// Mitsubishi GX Works2 project: TRANG TRAI   PLC: FX3U/FX3UC

PROGRAM MAIN
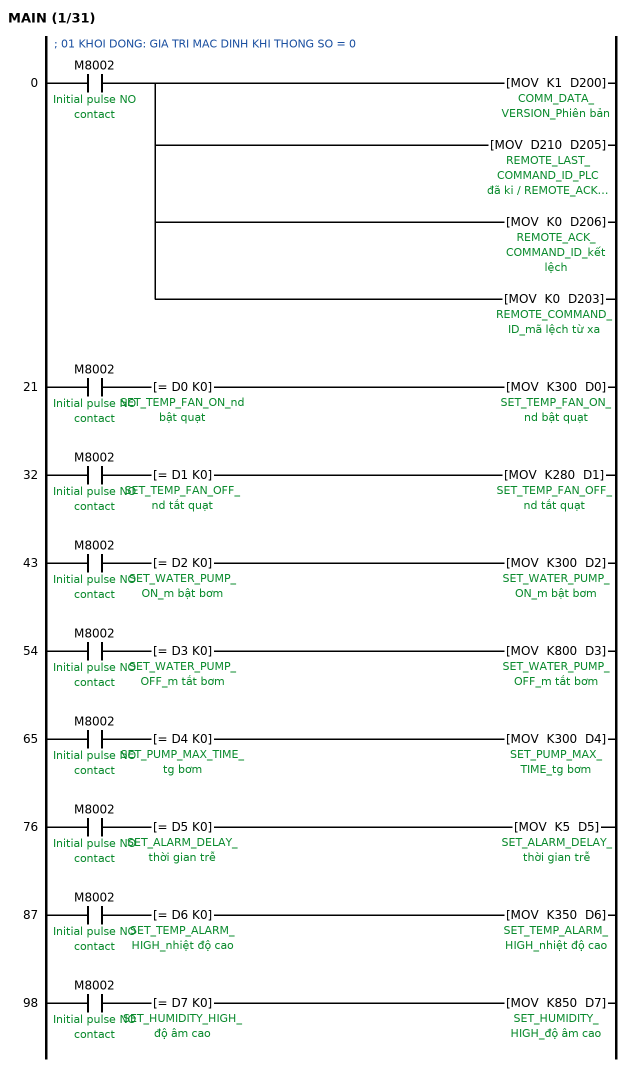
; 01 KHOI DONG: GIA TRI MAC DINH KHI THONG SO = 0
0     LD      M8002  ; Initial pulse NO contact
      MOV     K1 D200  ; COMM_DATA_VERSION_Phiên bản
      MOV     D210 D205  ; REMOTE_LAST_COMMAND_ID_PLC đã ki / REMOTE_ACK_COMMAND_ID_PLC đã nhậ
      MOV     K0 D206  ; REMOTE_ACK_COMMAND_ID_kết lệch
      MOV     K0 D203  ; REMOTE_COMMAND_ID_mã lệch từ xa
21    LD      M8002  ; Initial pulse NO contact
      AND=    D0 K0  ; SET_TEMP_FAN_ON_nd bật quạt
      MOV     K300 D0
32    LD      M8002  ; Initial pulse NO contact
      AND=    D1 K0  ; SET_TEMP_FAN_OFF_nd tắt quạt
      MOV     K280 D1
43    LD      M8002  ; Initial pulse NO contact
      AND=    D2 K0  ; SET_WATER_PUMP_ON_m bật bơm
      MOV     K300 D2
54    LD      M8002  ; Initial pulse NO contact
      AND=    D3 K0  ; SET_WATER_PUMP_OFF_m tắt bơm
      MOV     K800 D3
65    LD      M8002  ; Initial pulse NO contact
      AND=    D4 K0  ; SET_PUMP_MAX_TIME_tg bơm
      MOV     K300 D4
76    LD      M8002  ; Initial pulse NO contact
      AND=    D5 K0  ; SET_ALARM_DELAY_thời gian trễ
      MOV     K5 D5
87    LD      M8002  ; Initial pulse NO contact
      AND=    D6 K0  ; SET_TEMP_ALARM_HIGH_nhiệt độ cao
      MOV     K350 D6
98    LD      M8002  ; Initial pulse NO contact
      AND=    D7 K0  ; SET_HUMIDITY_HIGH_độ âm cao
      MOV     K850 D7
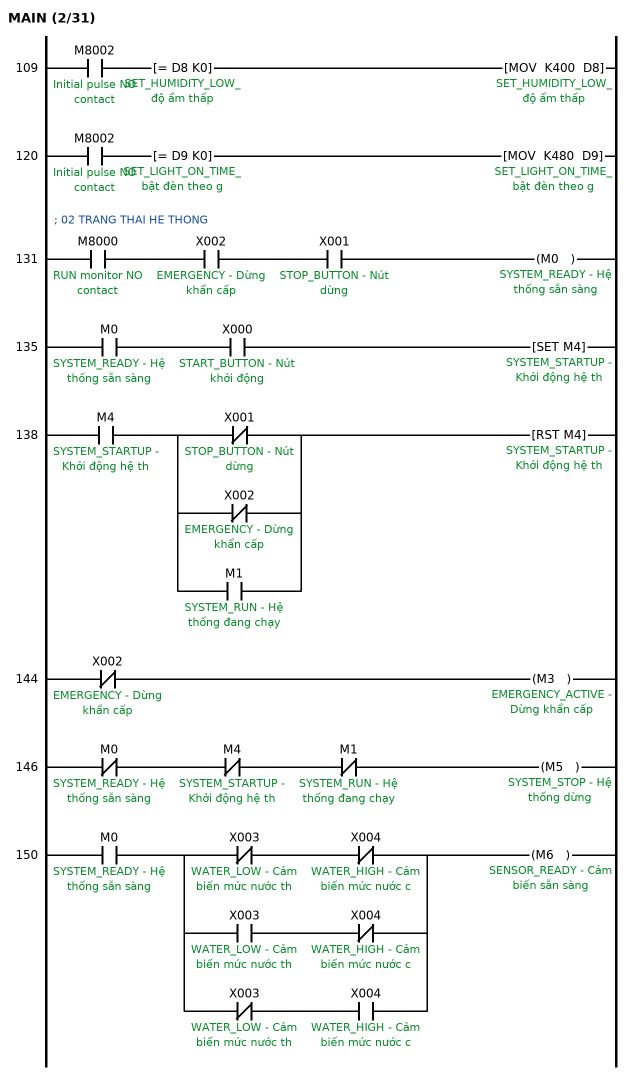
109   LD      M8002  ; Initial pulse NO contact
      AND=    D8 K0  ; SET_HUMIDITY_LOW_độ ẩm thấp
      MOV     K400 D8
120   LD      M8002  ; Initial pulse NO contact
      AND=    D9 K0  ; SET_LIGHT_ON_TIME_bật đèn theo g
      MOV     K480 D9
; 02 TRANG THAI HE THONG
131   LD      M8000  ; RUN monitor NO contact
      AND     X002  ; EMERGENCY - Dừng khẩn cấp
      AND     X001  ; STOP_BUTTON - Nút dừng
      OUT     M0  ; SYSTEM_READY - Hệ thống sẵn sàng
135   LD      M0  ; SYSTEM_READY - Hệ thống sẵn sàng
      AND     X000  ; START_BUTTON - Nút khởi động
      SET     M4  ; SYSTEM_STARTUP - Khởi động hệ th
138   LD      M4  ; SYSTEM_STARTUP - Khởi động hệ th
      LDI     X001  ; STOP_BUTTON - Nút dừng
      ORI     X002  ; EMERGENCY - Dừng khẩn cấp
      OR      M1  ; SYSTEM_RUN - Hệ thống đang chạy
      ANB
      RST     M4  ; SYSTEM_STARTUP - Khởi động hệ th
144   LDI     X002  ; EMERGENCY - Dừng khẩn cấp
      OUT     M3  ; EMERGENCY_ACTIVE - Dừng khẩn cấp
146   LDI     M0  ; SYSTEM_READY - Hệ thống sẵn sàng
      ANI     M4  ; SYSTEM_STARTUP - Khởi động hệ th
      ANI     M1  ; SYSTEM_RUN - Hệ thống đang chạy
      OUT     M5  ; SYSTEM_STOP - Hệ thống dừng
150   LD      M0  ; SYSTEM_READY - Hệ thống sẵn sàng
      LDI     X003  ; WATER_LOW - Cảm biến mức nước th
      ANI     X004  ; WATER_HIGH - Cảm biến mức nước c
      LD      X003  ; WATER_LOW - Cảm biến mức nước th
      ANI     X004  ; WATER_HIGH - Cảm biến mức nước c
      ORB
      LDI     X003  ; WATER_LOW - Cảm biến mức nước th
      AND     X004  ; WATER_HIGH - Cảm biến mức nước c
      ORB
      ANB
      OUT     M6  ; SENSOR_READY - Cảm biến sẵn sàng
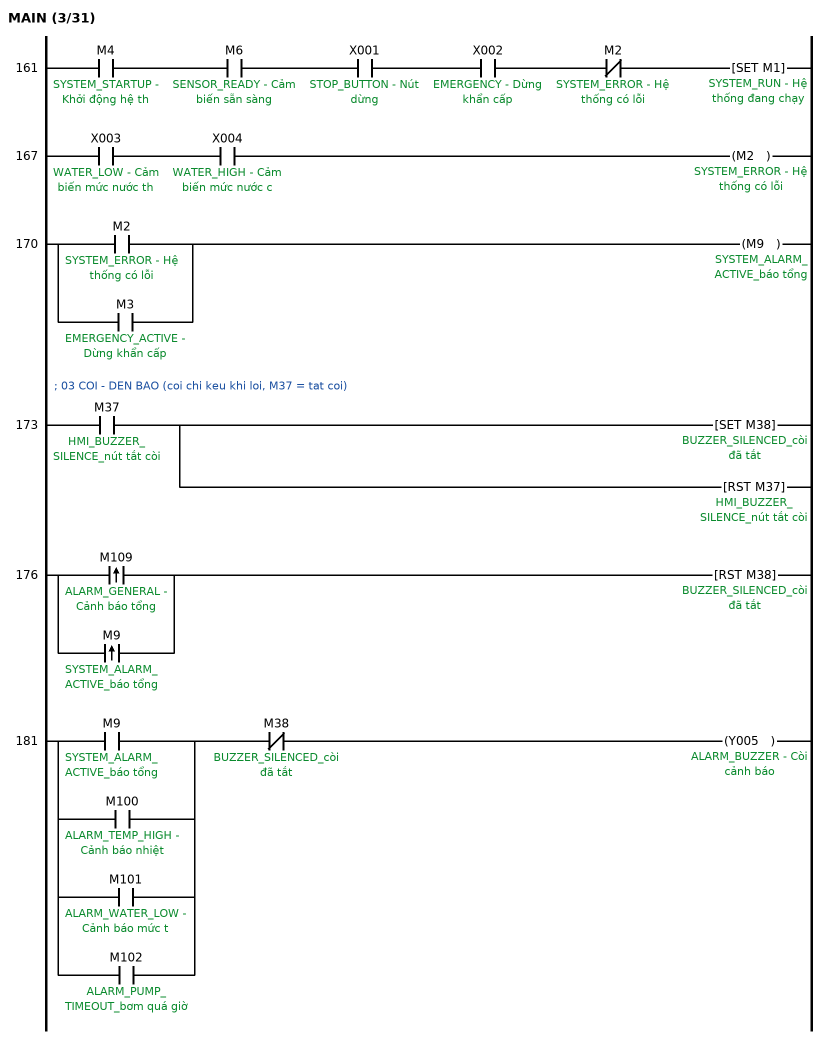
161   LD      M4  ; SYSTEM_STARTUP - Khởi động hệ th
      AND     M6  ; SENSOR_READY - Cảm biến sẵn sàng
      AND     X001  ; STOP_BUTTON - Nút dừng
      AND     X002  ; EMERGENCY - Dừng khẩn cấp
      ANI     M2  ; SYSTEM_ERROR - Hệ thống có lỗi
      SET     M1  ; SYSTEM_RUN - Hệ thống đang chạy
167   LD      X003  ; WATER_LOW - Cảm biến mức nước th
      AND     X004  ; WATER_HIGH - Cảm biến mức nước c
      OUT     M2  ; SYSTEM_ERROR - Hệ thống có lỗi
170   LD      M2  ; SYSTEM_ERROR - Hệ thống có lỗi
      OR      M3  ; EMERGENCY_ACTIVE - Dừng khẩn cấp
      OUT     M9  ; SYSTEM_ALARM_ACTIVE_báo tổng
; 03 COI - DEN BAO (coi chi keu khi loi, M37 = tat coi)
173   LD      M37  ; HMI_BUZZER_SILENCE_nút tắt còi
      SET     M38  ; BUZZER_SILENCED_còi đã tắt
      RST     M37  ; HMI_BUZZER_SILENCE_nút tắt còi
176   LDP     M109  ; ALARM_GENERAL - Cảnh báo tổng
      ORP     M9  ; SYSTEM_ALARM_ACTIVE_báo tổng
      RST     M38  ; BUZZER_SILENCED_còi đã tắt
181   LD      M9  ; SYSTEM_ALARM_ACTIVE_báo tổng
      OR      M100  ; ALARM_TEMP_HIGH - Cảnh báo nhiệt
      OR      M101  ; ALARM_WATER_LOW - Cảnh báo mức t
      OR      M102  ; ALARM_PUMP_TIMEOUT_bơm quá giờ
      ANI     M38  ; BUZZER_SILENCED_còi đã tắt
      OUT     Y005  ; ALARM_BUZZER - Còi cảnh báo
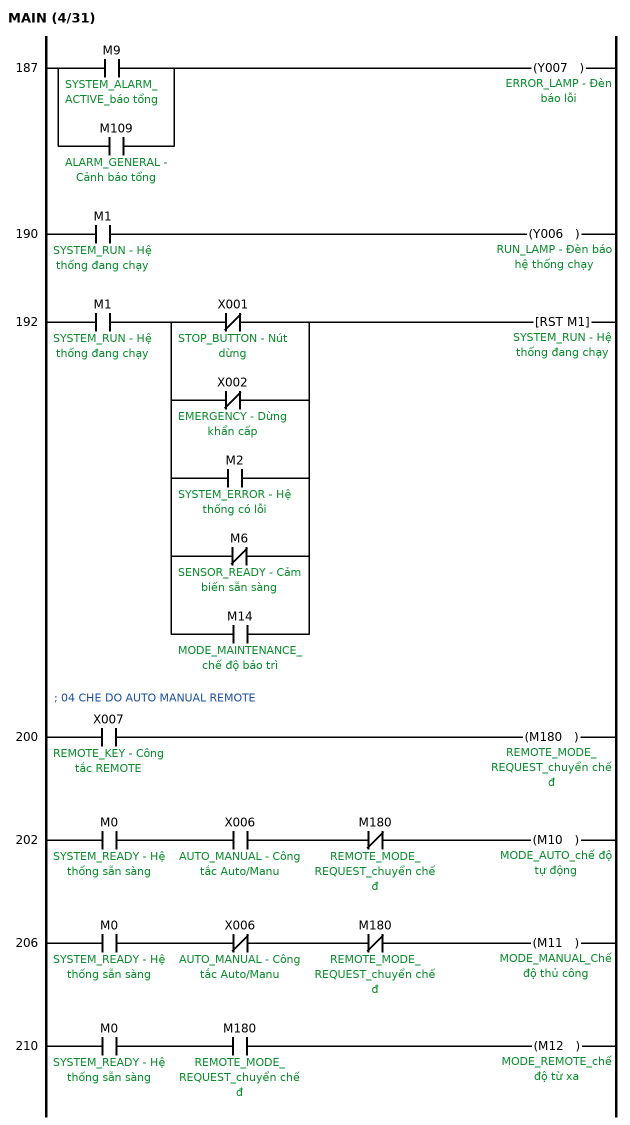
187   LD      M9  ; SYSTEM_ALARM_ACTIVE_báo tổng
      OR      M109  ; ALARM_GENERAL - Cảnh báo tổng
      OUT     Y007  ; ERROR_LAMP - Đèn báo lỗi
190   LD      M1  ; SYSTEM_RUN - Hệ thống đang chạy
      OUT     Y006  ; RUN_LAMP - Đèn báo hệ thống chạy
192   LD      M1  ; SYSTEM_RUN - Hệ thống đang chạy
      LDI     X001  ; STOP_BUTTON - Nút dừng
      ORI     X002  ; EMERGENCY - Dừng khẩn cấp
      OR      M2  ; SYSTEM_ERROR - Hệ thống có lỗi
      ORI     M6  ; SENSOR_READY - Cảm biến sẵn sàng
      OR      M14  ; MODE_MAINTENANCE_chế độ bảo trì
      ANB
      RST     M1  ; SYSTEM_RUN - Hệ thống đang chạy
; 04 CHE DO AUTO MANUAL REMOTE
200   LD      X007  ; REMOTE_KEY - Công tắc REMOTE
      OUT     M180  ; REMOTE_MODE_REQUEST_chuyển chế đ
202   LD      M0  ; SYSTEM_READY - Hệ thống sẵn sàng
      AND     X006  ; AUTO_MANUAL - Công tắc Auto/Manu
      ANI     M180  ; REMOTE_MODE_REQUEST_chuyển chế đ
      OUT     M10  ; MODE_AUTO_chế độ tự động
206   LD      M0  ; SYSTEM_READY - Hệ thống sẵn sàng
      ANI     X006  ; AUTO_MANUAL - Công tắc Auto/Manu
      ANI     M180  ; REMOTE_MODE_REQUEST_chuyển chế đ
      OUT     M11  ; MODE_MANUAL_Chế độ thủ công
210   LD      M0  ; SYSTEM_READY - Hệ thống sẵn sàng
      AND     M180  ; REMOTE_MODE_REQUEST_chuyển chế đ
      OUT     M12  ; MODE_REMOTE_chế độ từ xa
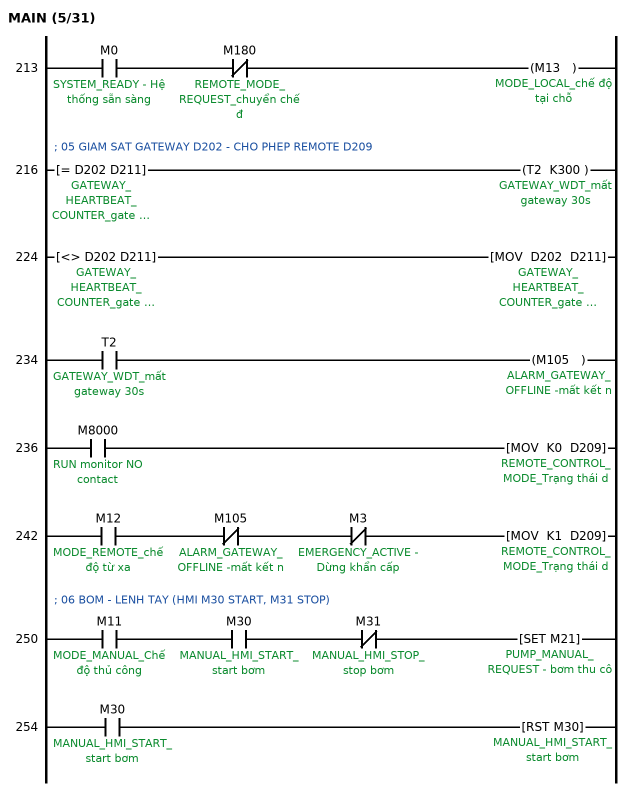
213   LD      M0  ; SYSTEM_READY - Hệ thống sẵn sàng
      ANI     M180  ; REMOTE_MODE_REQUEST_chuyển chế đ
      OUT     M13  ; MODE_LOCAL_chế độ tại chỗ
; 05 GIAM SAT GATEWAY D202 - CHO PHEP REMOTE D209
216   LD=     D202 D211  ; GATEWAY_HEARTBEAT_COUNTER_gate / GATEWAY_HB_LAST_D202 lần trước
      OUT     T2 K300  ; GATEWAY_WDT_mất gateway 30s
224   LD<>    D202 D211  ; GATEWAY_HEARTBEAT_COUNTER_gate / GATEWAY_HB_LAST_D202 lần trước
      MOV     D202 D211
234   LD      T2  ; GATEWAY_WDT_mất gateway 30s
      OUT     M105  ; ALARM_GATEWAY_OFFLINE -mất kết n
236   LD      M8000  ; RUN monitor NO contact
      MOV     K0 D209  ; REMOTE_CONTROL_MODE_Trạng thái d
242   LD      M12  ; MODE_REMOTE_chế độ từ xa
      ANI     M105  ; ALARM_GATEWAY_OFFLINE -mất kết n
      ANI     M3  ; EMERGENCY_ACTIVE - Dừng khẩn cấp
      MOV     K1 D209
; 06 BOM - LENH TAY (HMI M30 START, M31 STOP)
250   LD      M11  ; MODE_MANUAL_Chế độ thủ công
      AND     M30  ; MANUAL_HMI_START_start bơm
      ANI     M31  ; MANUAL_HMI_STOP_stop bơm
      SET     M21  ; PUMP_MANUAL_REQUEST - bơm thu cô
254   LD      M30  ; MANUAL_HMI_START_start bơm
      RST     M30  ; MANUAL_HMI_START_start bơm
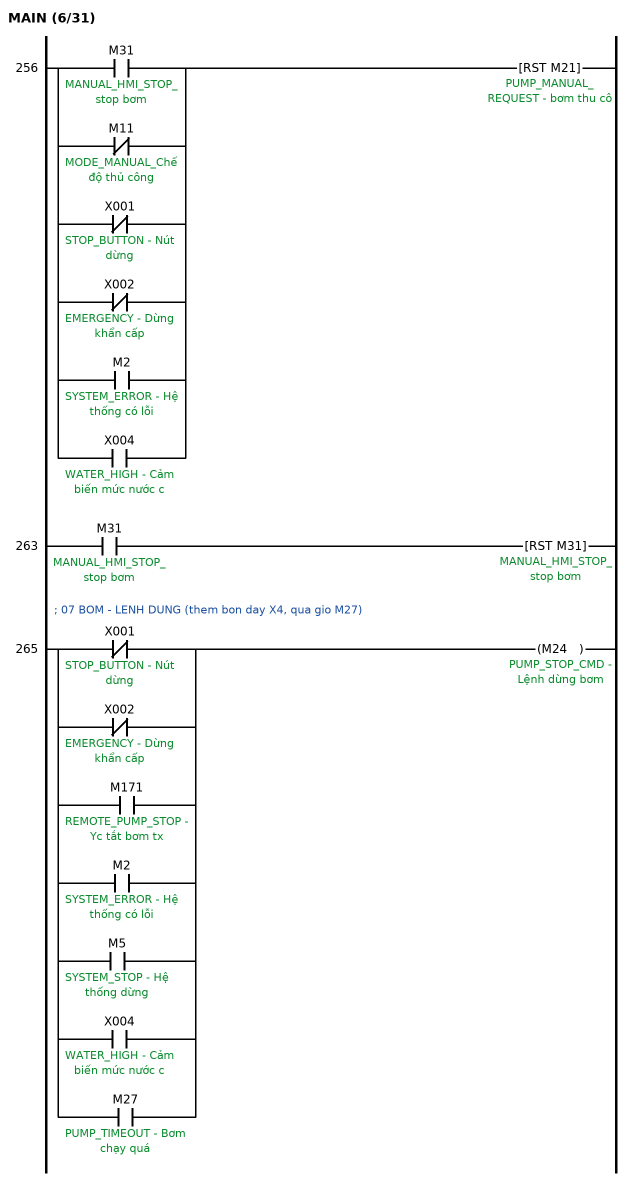
256   LD      M31  ; MANUAL_HMI_STOP_stop bơm
      ORI     M11  ; MODE_MANUAL_Chế độ thủ công
      ORI     X001  ; STOP_BUTTON - Nút dừng
      ORI     X002  ; EMERGENCY - Dừng khẩn cấp
      OR      M2  ; SYSTEM_ERROR - Hệ thống có lỗi
      OR      X004  ; WATER_HIGH - Cảm biến mức nước c
      RST     M21  ; PUMP_MANUAL_REQUEST - bơm thu cô
263   LD      M31  ; MANUAL_HMI_STOP_stop bơm
      RST     M31  ; MANUAL_HMI_STOP_stop bơm
; 07 BOM - LENH DUNG (them bon day X4, qua gio M27)
265   LDI     X001  ; STOP_BUTTON - Nút dừng
      ORI     X002  ; EMERGENCY - Dừng khẩn cấp
      OR      M171  ; REMOTE_PUMP_STOP - Yc tắt bơm tx
      OR      M2  ; SYSTEM_ERROR - Hệ thống có lỗi
      OR      M5  ; SYSTEM_STOP - Hệ thống dừng
      OR      X004  ; WATER_HIGH - Cảm biến mức nước c
      OR      M27  ; PUMP_TIMEOUT - Bơm chạy quá
      OUT     M24  ; PUMP_STOP_CMD - Lệnh dừng bơm
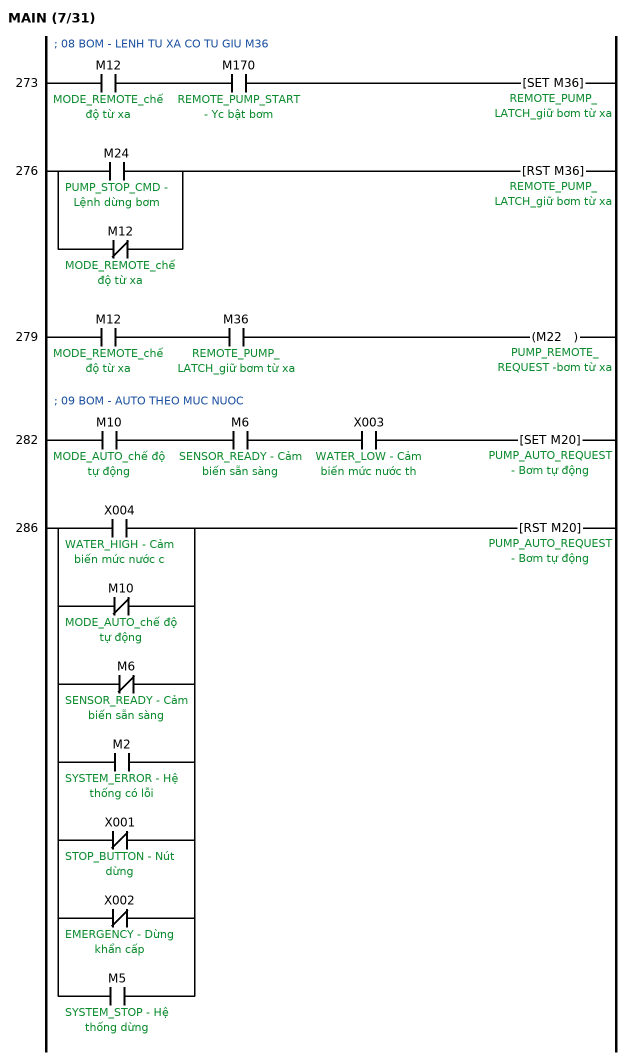
; 08 BOM - LENH TU XA CO TU GIU M36
273   LD      M12  ; MODE_REMOTE_chế độ từ xa
      AND     M170  ; REMOTE_PUMP_START - Yc bật bơm
      SET     M36  ; REMOTE_PUMP_LATCH_giữ bơm từ xa
276   LD      M24  ; PUMP_STOP_CMD - Lệnh dừng bơm
      ORI     M12  ; MODE_REMOTE_chế độ từ xa
      RST     M36  ; REMOTE_PUMP_LATCH_giữ bơm từ xa
279   LD      M12  ; MODE_REMOTE_chế độ từ xa
      AND     M36  ; REMOTE_PUMP_LATCH_giữ bơm từ xa
      OUT     M22  ; PUMP_REMOTE_REQUEST -bơm từ xa
; 09 BOM - AUTO THEO MUC NUOC
282   LD      M10  ; MODE_AUTO_chế độ tự động
      AND     M6  ; SENSOR_READY - Cảm biến sẵn sàng
      AND     X003  ; WATER_LOW - Cảm biến mức nước th
      SET     M20  ; PUMP_AUTO_REQUEST - Bơm tự động
286   LD      X004  ; WATER_HIGH - Cảm biến mức nước c
      ORI     M10  ; MODE_AUTO_chế độ tự động
      ORI     M6  ; SENSOR_READY - Cảm biến sẵn sàng
      OR      M2  ; SYSTEM_ERROR - Hệ thống có lỗi
      ORI     X001  ; STOP_BUTTON - Nút dừng
      ORI     X002  ; EMERGENCY - Dừng khẩn cấp
      OR      M5  ; SYSTEM_STOP - Hệ thống dừng
      RST     M20  ; PUMP_AUTO_REQUEST - Bơm tự động
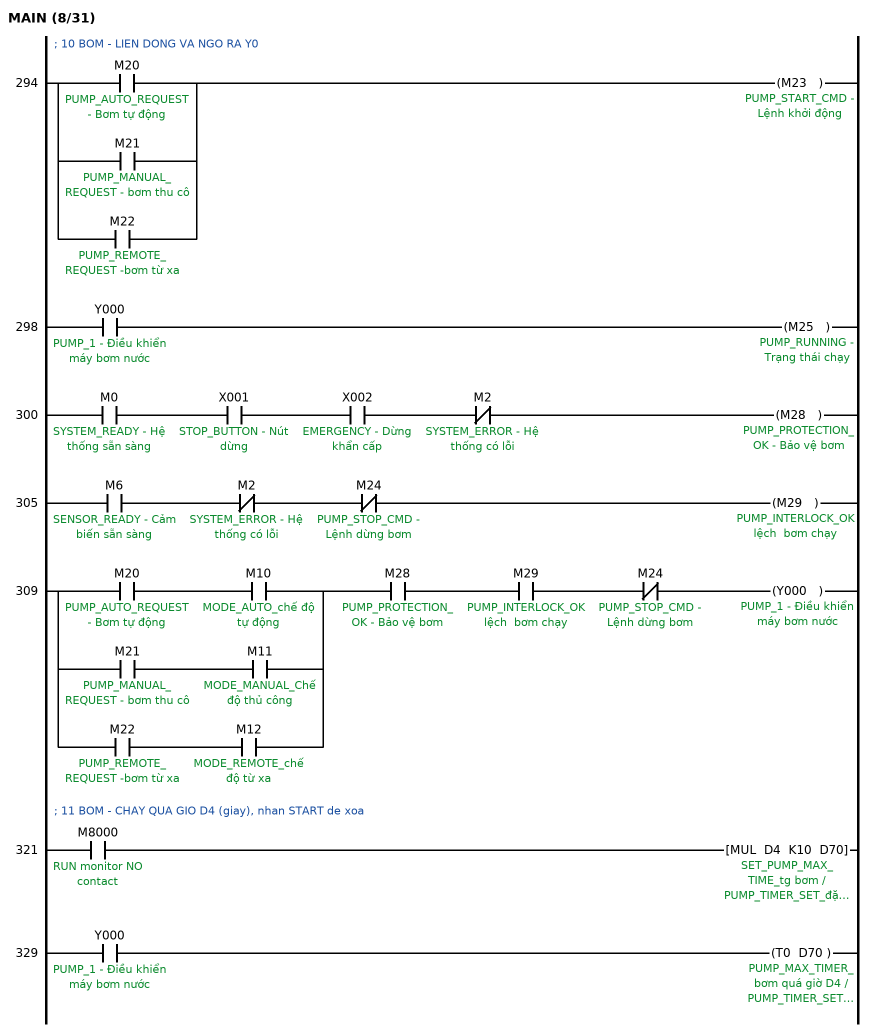
; 10 BOM - LIEN DONG VA NGO RA Y0
294   LD      M20  ; PUMP_AUTO_REQUEST - Bơm tự động
      OR      M21  ; PUMP_MANUAL_REQUEST - bơm thu cô
      OR      M22  ; PUMP_REMOTE_REQUEST -bơm từ xa
      OUT     M23  ; PUMP_START_CMD - Lệnh khởi động
298   LD      Y000  ; PUMP_1 - Điều khiển máy bơm nước
      OUT     M25  ; PUMP_RUNNING - Trạng thái chạy
300   LD      M0  ; SYSTEM_READY - Hệ thống sẵn sàng
      AND     X001  ; STOP_BUTTON - Nút dừng
      AND     X002  ; EMERGENCY - Dừng khẩn cấp
      ANI     M2  ; SYSTEM_ERROR - Hệ thống có lỗi
      OUT     M28  ; PUMP_PROTECTION_OK - Bảo vệ bơm
305   LD      M6  ; SENSOR_READY - Cảm biến sẵn sàng
      ANI     M2  ; SYSTEM_ERROR - Hệ thống có lỗi
      ANI     M24  ; PUMP_STOP_CMD - Lệnh dừng bơm
      OUT     M29  ; PUMP_INTERLOCK_OK lệch  bơm chạy
309   LD      M20  ; PUMP_AUTO_REQUEST - Bơm tự động
      AND     M10  ; MODE_AUTO_chế độ tự động
      LD      M21  ; PUMP_MANUAL_REQUEST - bơm thu cô
      AND     M11  ; MODE_MANUAL_Chế độ thủ công
      ORB
      LD      M22  ; PUMP_REMOTE_REQUEST -bơm từ xa
      AND     M12  ; MODE_REMOTE_chế độ từ xa
      ORB
      AND     M28  ; PUMP_PROTECTION_OK - Bảo vệ bơm
      AND     M29  ; PUMP_INTERLOCK_OK lệch  bơm chạy
      ANI     M24  ; PUMP_STOP_CMD - Lệnh dừng bơm
      OUT     Y000  ; PUMP_1 - Điều khiển máy bơm nước
; 11 BOM - CHAY QUA GIO D4 (giay), nhan START de xoa
321   LD      M8000  ; RUN monitor NO contact
      MUL     D4 K10 D70  ; PUMP_TIMER_SET_đặt T0 = D4x10
329   LD      Y000  ; PUMP_1 - Điều khiển máy bơm nước
      OUT     T0 D70  ; PUMP_MAX_TIMER_bơm quá giờ D4 / PUMP_TIMER_SET_đặt T0 = D4x10
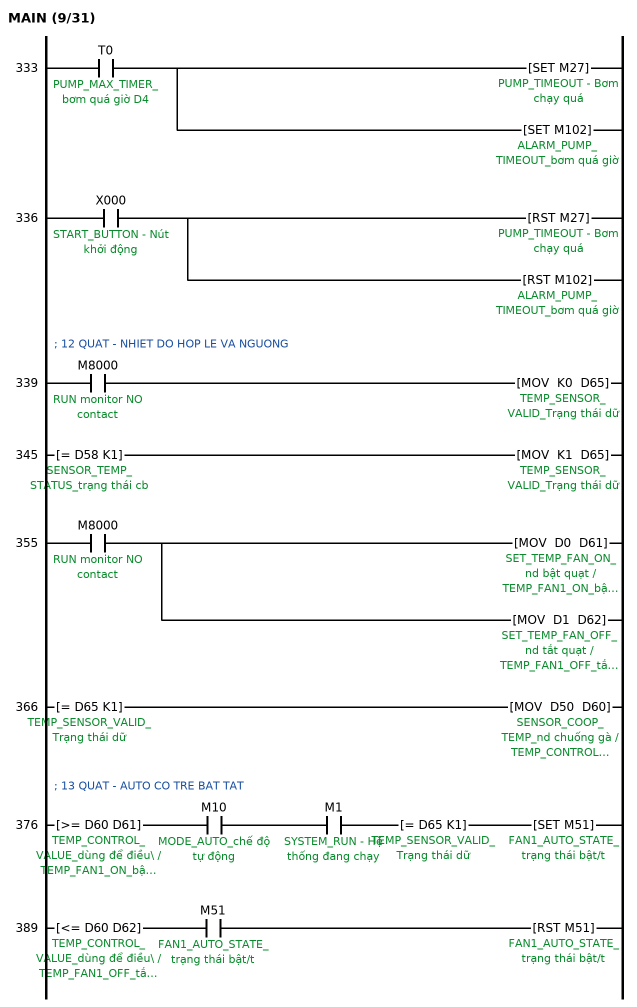
333   LD      T0  ; PUMP_MAX_TIMER_bơm quá giờ D4
      SET     M27  ; PUMP_TIMEOUT - Bơm chạy quá
      SET     M102  ; ALARM_PUMP_TIMEOUT_bơm quá giờ
336   LD      X000  ; START_BUTTON - Nút khởi động
      RST     M27  ; PUMP_TIMEOUT - Bơm chạy quá
      RST     M102  ; ALARM_PUMP_TIMEOUT_bơm quá giờ
; 12 QUAT - NHIET DO HOP LE VA NGUONG
339   LD      M8000  ; RUN monitor NO contact
      MOV     K0 D65  ; TEMP_SENSOR_VALID_Trạng thái dữ
345   LD=     D58 K1  ; SENSOR_TEMP_STATUS_trạng thái cb
      MOV     K1 D65
355   LD      M8000  ; RUN monitor NO contact
      MOV     D0 D61  ; TEMP_FAN1_ON_bật quạt 1
      MOV     D1 D62  ; TEMP_FAN1_OFF_tắt quạt 1
366   LD=     D65 K1  ; TEMP_SENSOR_VALID_Trạng thái dữ
      MOV     D50 D60  ; SENSOR_COOP_TEMP_nd chuống gà / TEMP_CONTROL_VALUE_dùng để điều\
; 13 QUAT - AUTO CO TRE BAT TAT
376   LD>=    D60 D61  ; TEMP_CONTROL_VALUE_dùng để điều\ / TEMP_FAN1_ON_bật quạt 1
      AND     M10  ; MODE_AUTO_chế độ tự động
      AND     M1  ; SYSTEM_RUN - Hệ thống đang chạy
      AND=    D65 K1  ; TEMP_SENSOR_VALID_Trạng thái dữ
      SET     M51  ; FAN1_AUTO_STATE_trạng thái bật/t
389   LD<=    D60 D62  ; TEMP_CONTROL_VALUE_dùng để điều\ / TEMP_FAN1_OFF_tắt quạt 1
      AND     M51  ; FAN1_AUTO_STATE_trạng thái bật/t
      RST     M51  ; FAN1_AUTO_STATE_trạng thái bật/t
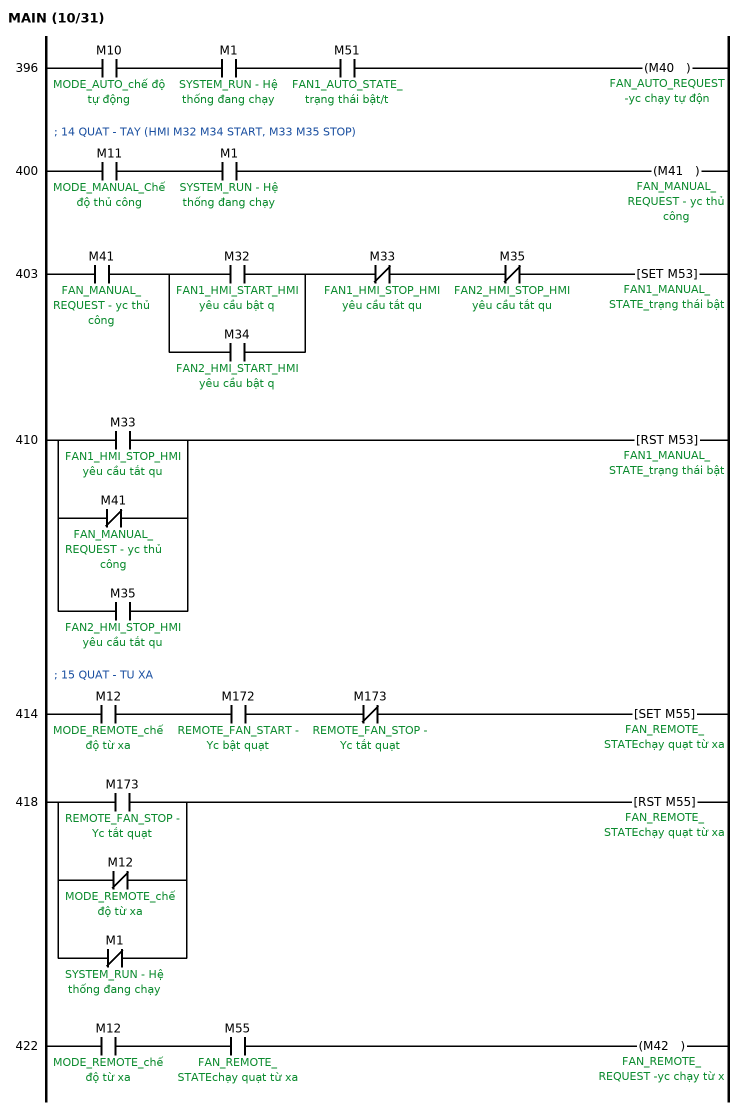
396   LD      M10  ; MODE_AUTO_chế độ tự động
      AND     M1  ; SYSTEM_RUN - Hệ thống đang chạy
      AND     M51  ; FAN1_AUTO_STATE_trạng thái bật/t
      OUT     M40  ; FAN_AUTO_REQUEST -yc chạy tự độn
; 14 QUAT - TAY (HMI M32 M34 START, M33 M35 STOP)
400   LD      M11  ; MODE_MANUAL_Chế độ thủ công
      AND     M1  ; SYSTEM_RUN - Hệ thống đang chạy
      OUT     M41  ; FAN_MANUAL_REQUEST - yc thủ công
403   LD      M41  ; FAN_MANUAL_REQUEST - yc thủ công
      LD      M32  ; FAN1_HMI_START_HMI yêu cầu bật q
      OR      M34  ; FAN2_HMI_START_HMI yêu cầu bật q
      ANB
      ANI     M33  ; FAN1_HMI_STOP_HMI yêu cầu tắt qu
      ANI     M35  ; FAN2_HMI_STOP_HMI yêu cầu tắt qu
      SET     M53  ; FAN1_MANUAL_STATE_trạng thái bật
410   LD      M33  ; FAN1_HMI_STOP_HMI yêu cầu tắt qu
      ORI     M41  ; FAN_MANUAL_REQUEST - yc thủ công
      OR      M35  ; FAN2_HMI_STOP_HMI yêu cầu tắt qu
      RST     M53  ; FAN1_MANUAL_STATE_trạng thái bật
; 15 QUAT - TU XA
414   LD      M12  ; MODE_REMOTE_chế độ từ xa
      AND     M172  ; REMOTE_FAN_START - Yc bật quạt
      ANI     M173  ; REMOTE_FAN_STOP - Yc tắt quạt
      SET     M55  ; FAN_REMOTE_STATEchạy quạt từ xa
418   LD      M173  ; REMOTE_FAN_STOP - Yc tắt quạt
      ORI     M12  ; MODE_REMOTE_chế độ từ xa
      ORI     M1  ; SYSTEM_RUN - Hệ thống đang chạy
      RST     M55  ; FAN_REMOTE_STATEchạy quạt từ xa
422   LD      M12  ; MODE_REMOTE_chế độ từ xa
      AND     M55  ; FAN_REMOTE_STATEchạy quạt từ xa
      OUT     M42  ; FAN_REMOTE_REQUEST -yc chạy từ x
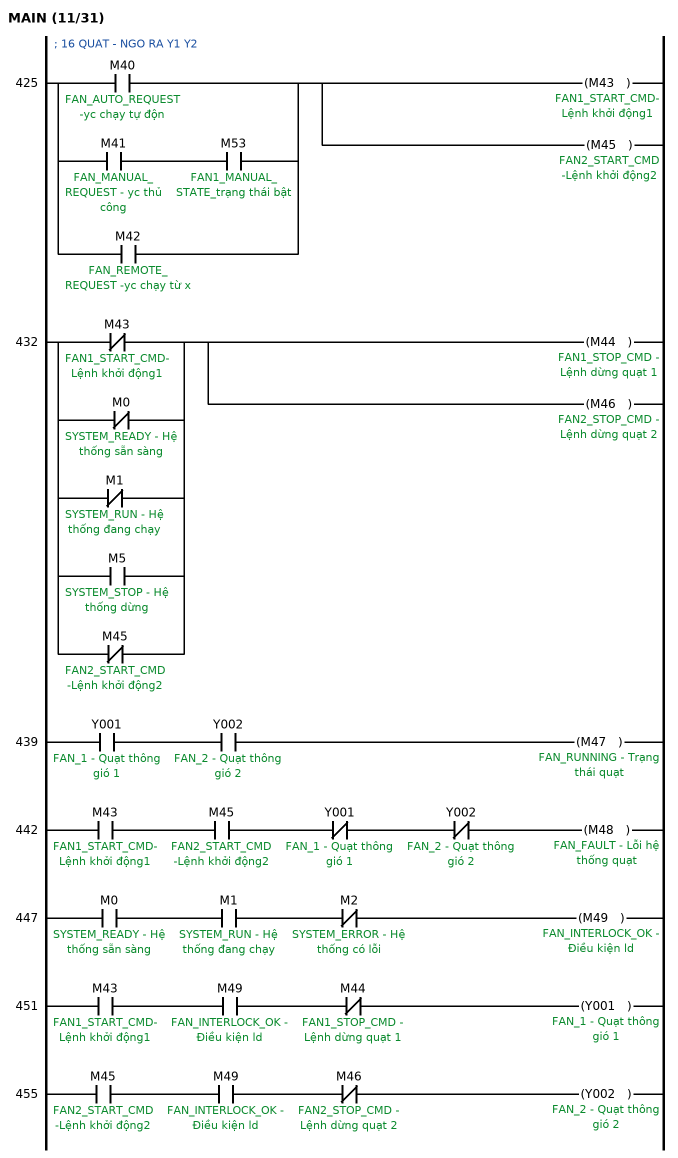
; 16 QUAT - NGO RA Y1 Y2
425   LD      M40  ; FAN_AUTO_REQUEST -yc chạy tự độn
      LD      M41  ; FAN_MANUAL_REQUEST - yc thủ công
      AND     M53  ; FAN1_MANUAL_STATE_trạng thái bật
      ORB
      OR      M42  ; FAN_REMOTE_REQUEST -yc chạy từ x
      OUT     M43  ; FAN1_START_CMD-Lệnh khởi động1
      OUT     M45  ; FAN2_START_CMD -Lệnh khởi động2
432   LDI     M43  ; FAN1_START_CMD-Lệnh khởi động1
      ORI     M0  ; SYSTEM_READY - Hệ thống sẵn sàng
      ORI     M1  ; SYSTEM_RUN - Hệ thống đang chạy
      OR      M5  ; SYSTEM_STOP - Hệ thống dừng
      ORI     M45  ; FAN2_START_CMD -Lệnh khởi động2
      OUT     M44  ; FAN1_STOP_CMD - Lệnh dừng quạt 1
      OUT     M46  ; FAN2_STOP_CMD - Lệnh dừng quạt 2
439   LD      Y001  ; FAN_1 - Quạt thông gió 1
      AND     Y002  ; FAN_2 - Quạt thông gió 2
      OUT     M47  ; FAN_RUNNING - Trạng thái quạt
442   LD      M43  ; FAN1_START_CMD-Lệnh khởi động1
      AND     M45  ; FAN2_START_CMD -Lệnh khởi động2
      ANI     Y001  ; FAN_1 - Quạt thông gió 1
      ANI     Y002  ; FAN_2 - Quạt thông gió 2
      OUT     M48  ; FAN_FAULT - Lỗi hệ thống quạt
447   LD      M0  ; SYSTEM_READY - Hệ thống sẵn sàng
      AND     M1  ; SYSTEM_RUN - Hệ thống đang chạy
      ANI     M2  ; SYSTEM_ERROR - Hệ thống có lỗi
      OUT     M49  ; FAN_INTERLOCK_OK - Điều kiện ld
451   LD      M43  ; FAN1_START_CMD-Lệnh khởi động1
      AND     M49  ; FAN_INTERLOCK_OK - Điều kiện ld
      ANI     M44  ; FAN1_STOP_CMD - Lệnh dừng quạt 1
      OUT     Y001  ; FAN_1 - Quạt thông gió 1
455   LD      M45  ; FAN2_START_CMD -Lệnh khởi động2
      AND     M49  ; FAN_INTERLOCK_OK - Điều kiện ld
      ANI     M46  ; FAN2_STOP_CMD - Lệnh dừng quạt 2
      OUT     Y002  ; FAN_2 - Quạt thông gió 2
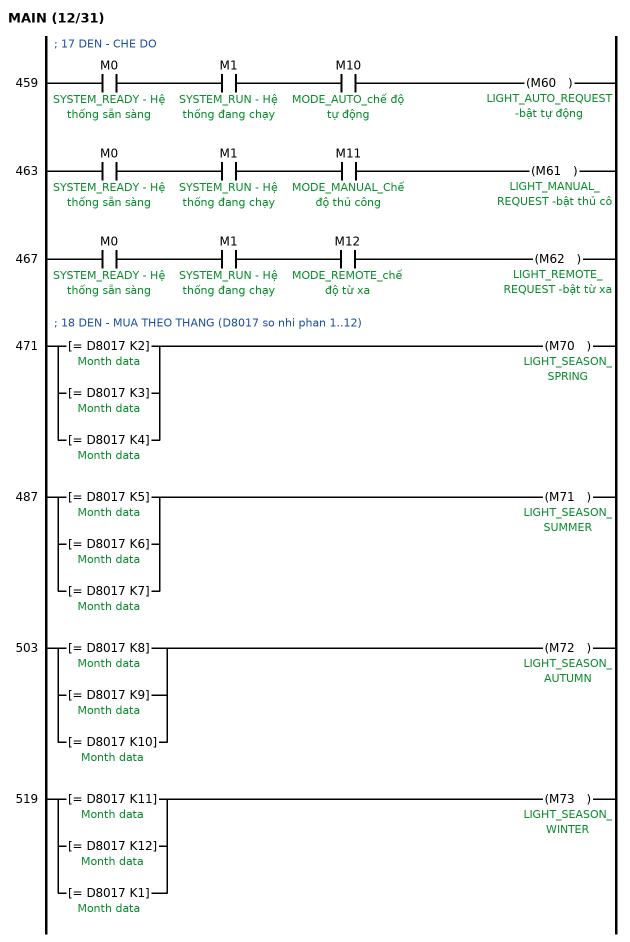
; 17 DEN - CHE DO
459   LD      M0  ; SYSTEM_READY - Hệ thống sẵn sàng
      AND     M1  ; SYSTEM_RUN - Hệ thống đang chạy
      AND     M10  ; MODE_AUTO_chế độ tự động
      OUT     M60  ; LIGHT_AUTO_REQUEST -bật tự động
463   LD      M0  ; SYSTEM_READY - Hệ thống sẵn sàng
      AND     M1  ; SYSTEM_RUN - Hệ thống đang chạy
      AND     M11  ; MODE_MANUAL_Chế độ thủ công
      OUT     M61  ; LIGHT_MANUAL_REQUEST -bật thủ cô
467   LD      M0  ; SYSTEM_READY - Hệ thống sẵn sàng
      AND     M1  ; SYSTEM_RUN - Hệ thống đang chạy
      AND     M12  ; MODE_REMOTE_chế độ từ xa
      OUT     M62  ; LIGHT_REMOTE_REQUEST -bật từ xa
; 18 DEN - MUA THEO THANG (D8017 so nhi phan 1..12)
471   LD=     D8017 K2  ; Month data
      OR=     D8017 K3  ; Month data
      OR=     D8017 K4  ; Month data
      OUT     M70  ; LIGHT_SEASON_SPRING
487   LD=     D8017 K5  ; Month data
      OR=     D8017 K6  ; Month data
      OR=     D8017 K7  ; Month data
      OUT     M71  ; LIGHT_SEASON_SUMMER
503   LD=     D8017 K8  ; Month data
      OR=     D8017 K9  ; Month data
      OR=     D8017 K10  ; Month data
      OUT     M72  ; LIGHT_SEASON_AUTUMN
519   LD=     D8017 K11  ; Month data
      OR=     D8017 K12  ; Month data
      OR=     D8017 K1  ; Month data
      OUT     M73  ; LIGHT_SEASON_WINTER
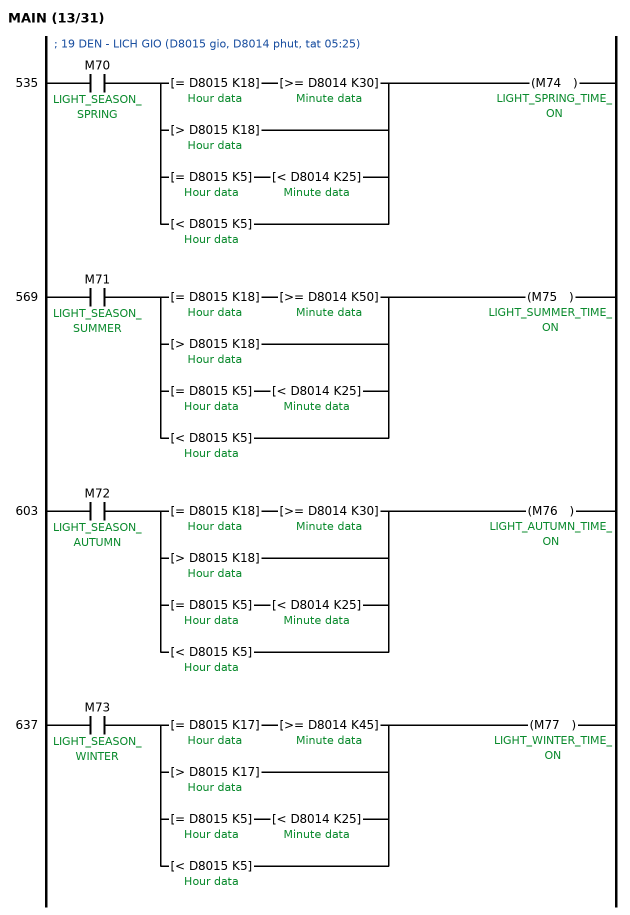
; 19 DEN - LICH GIO (D8015 gio, D8014 phut, tat 05:25)
535   LD      M70  ; LIGHT_SEASON_SPRING
      LD=     D8015 K18  ; Hour data
      AND>=   D8014 K30  ; Minute data
      OR>     D8015 K18  ; Hour data
      LD=     D8015 K5  ; Hour data
      AND<    D8014 K25  ; Minute data
      ORB
      OR<     D8015 K5  ; Hour data
      ANB
      OUT     M74  ; LIGHT_SPRING_TIME_ON
569   LD      M71  ; LIGHT_SEASON_SUMMER
      LD=     D8015 K18  ; Hour data
      AND>=   D8014 K50  ; Minute data
      OR>     D8015 K18  ; Hour data
      LD=     D8015 K5  ; Hour data
      AND<    D8014 K25  ; Minute data
      ORB
      OR<     D8015 K5  ; Hour data
      ANB
      OUT     M75  ; LIGHT_SUMMER_TIME_ON
603   LD      M72  ; LIGHT_SEASON_AUTUMN
      LD=     D8015 K18  ; Hour data
      AND>=   D8014 K30  ; Minute data
      OR>     D8015 K18  ; Hour data
      LD=     D8015 K5  ; Hour data
      AND<    D8014 K25  ; Minute data
      ORB
      OR<     D8015 K5  ; Hour data
      ANB
      OUT     M76  ; LIGHT_AUTUMN_TIME_ON
637   LD      M73  ; LIGHT_SEASON_WINTER
      LD=     D8015 K17  ; Hour data
      AND>=   D8014 K45  ; Minute data
      OR>     D8015 K17  ; Hour data
      LD=     D8015 K5  ; Hour data
      AND<    D8014 K25  ; Minute data
      ORB
      OR<     D8015 K5  ; Hour data
      ANB
      OUT     M77  ; LIGHT_WINTER_TIME_ON
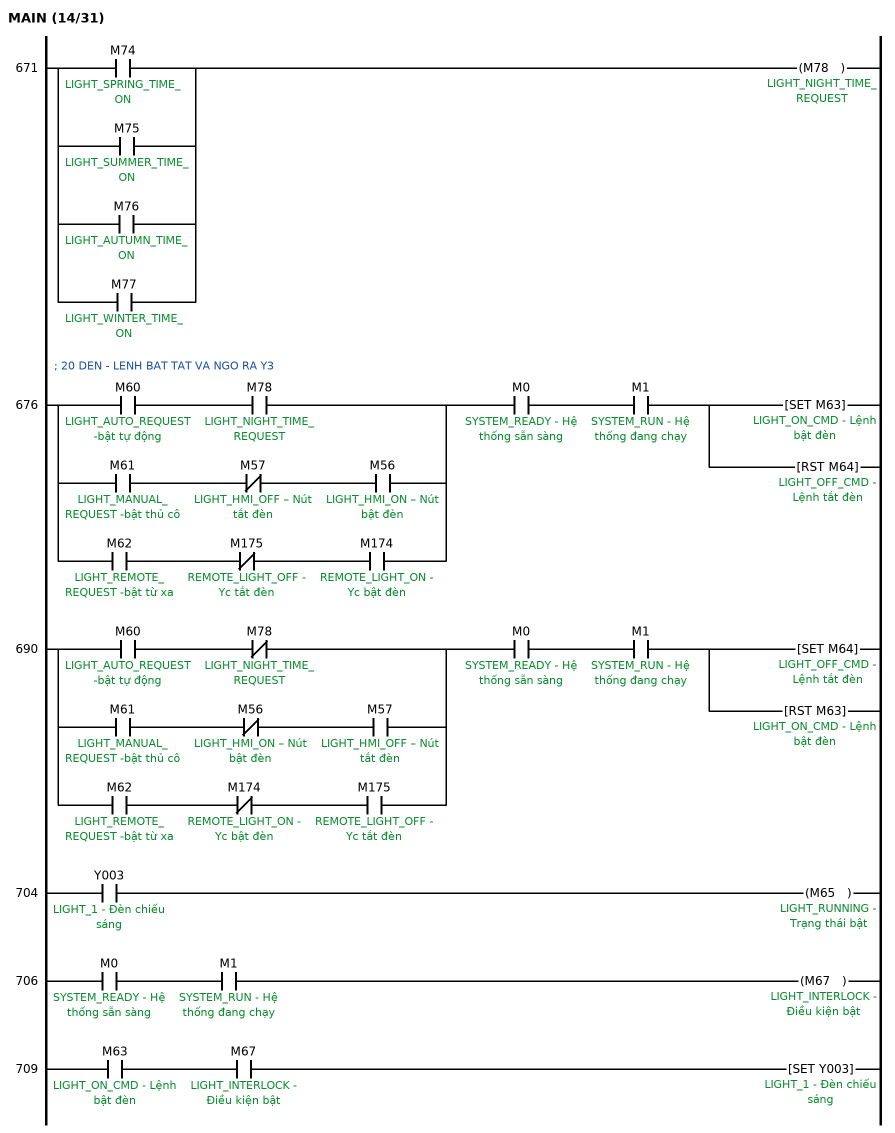
671   LD      M74  ; LIGHT_SPRING_TIME_ON
      OR      M75  ; LIGHT_SUMMER_TIME_ON
      OR      M76  ; LIGHT_AUTUMN_TIME_ON
      OR      M77  ; LIGHT_WINTER_TIME_ON
      OUT     M78  ; LIGHT_NIGHT_TIME_REQUEST
; 20 DEN - LENH BAT TAT VA NGO RA Y3
676   LD      M60  ; LIGHT_AUTO_REQUEST -bật tự động
      AND     M78  ; LIGHT_NIGHT_TIME_REQUEST
      LD      M61  ; LIGHT_MANUAL_REQUEST -bật thủ cô
      ANI     M57  ; LIGHT_HMI_OFF – Nút tắt đèn
      AND     M56  ; LIGHT_HMI_ON – Nút bật đèn
      ORB
      LD      M62  ; LIGHT_REMOTE_REQUEST -bật từ xa
      ANI     M175  ; REMOTE_LIGHT_OFF - Yc tắt đèn
      AND     M174  ; REMOTE_LIGHT_ON - Yc bật đèn
      ORB
      AND     M0  ; SYSTEM_READY - Hệ thống sẵn sàng
      AND     M1  ; SYSTEM_RUN - Hệ thống đang chạy
      SET     M63  ; LIGHT_ON_CMD - Lệnh bật đèn
      RST     M64  ; LIGHT_OFF_CMD - Lệnh tắt đèn
690   LD      M60  ; LIGHT_AUTO_REQUEST -bật tự động
      ANI     M78  ; LIGHT_NIGHT_TIME_REQUEST
      LD      M61  ; LIGHT_MANUAL_REQUEST -bật thủ cô
      ANI     M56  ; LIGHT_HMI_ON – Nút bật đèn
      AND     M57  ; LIGHT_HMI_OFF – Nút tắt đèn
      ORB
      LD      M62  ; LIGHT_REMOTE_REQUEST -bật từ xa
      ANI     M174  ; REMOTE_LIGHT_ON - Yc bật đèn
      AND     M175  ; REMOTE_LIGHT_OFF - Yc tắt đèn
      ORB
      AND     M0  ; SYSTEM_READY - Hệ thống sẵn sàng
      AND     M1  ; SYSTEM_RUN - Hệ thống đang chạy
      SET     M64  ; LIGHT_OFF_CMD - Lệnh tắt đèn
      RST     M63  ; LIGHT_ON_CMD - Lệnh bật đèn
704   LD      Y003  ; LIGHT_1 - Đèn chiếu sáng
      OUT     M65  ; LIGHT_RUNNING - Trạng thái bật
706   LD      M0  ; SYSTEM_READY - Hệ thống sẵn sàng
      AND     M1  ; SYSTEM_RUN - Hệ thống đang chạy
      OUT     M67  ; LIGHT_INTERLOCK - Điều kiện bật
709   LD      M63  ; LIGHT_ON_CMD - Lệnh bật đèn
      AND     M67  ; LIGHT_INTERLOCK - Điều kiện bật
      SET     Y003  ; LIGHT_1 - Đèn chiếu sáng
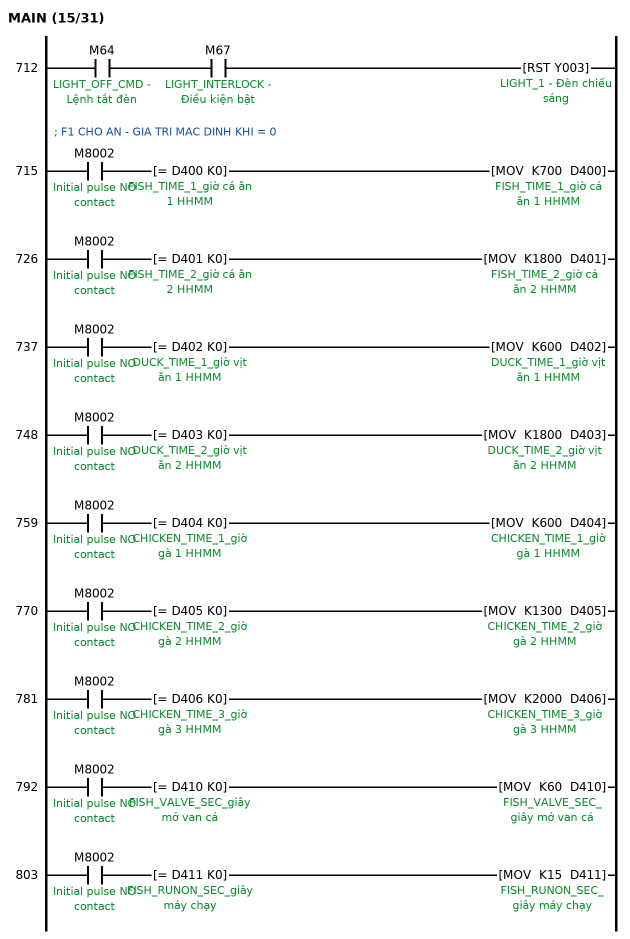
712   LD      M64  ; LIGHT_OFF_CMD - Lệnh tắt đèn
      AND     M67  ; LIGHT_INTERLOCK - Điều kiện bật
      RST     Y003  ; LIGHT_1 - Đèn chiếu sáng
; F1 CHO AN - GIA TRI MAC DINH KHI = 0
715   LD      M8002  ; Initial pulse NO contact
      AND=    D400 K0  ; FISH_TIME_1_giờ cá ăn 1 HHMM
      MOV     K700 D400
726   LD      M8002  ; Initial pulse NO contact
      AND=    D401 K0  ; FISH_TIME_2_giờ cá ăn 2 HHMM
      MOV     K1800 D401
737   LD      M8002  ; Initial pulse NO contact
      AND=    D402 K0  ; DUCK_TIME_1_giờ vịt ăn 1 HHMM
      MOV     K600 D402
748   LD      M8002  ; Initial pulse NO contact
      AND=    D403 K0  ; DUCK_TIME_2_giờ vịt ăn 2 HHMM
      MOV     K1800 D403
759   LD      M8002  ; Initial pulse NO contact
      AND=    D404 K0  ; CHICKEN_TIME_1_giờ gà 1 HHMM
      MOV     K600 D404
770   LD      M8002  ; Initial pulse NO contact
      AND=    D405 K0  ; CHICKEN_TIME_2_giờ gà 2 HHMM
      MOV     K1300 D405
781   LD      M8002  ; Initial pulse NO contact
      AND=    D406 K0  ; CHICKEN_TIME_3_giờ gà 3 HHMM
      MOV     K2000 D406
792   LD      M8002  ; Initial pulse NO contact
      AND=    D410 K0  ; FISH_VALVE_SEC_giây mở van cá
      MOV     K60 D410
803   LD      M8002  ; Initial pulse NO contact
      AND=    D411 K0  ; FISH_RUNON_SEC_giây máy chạy
      MOV     K15 D411
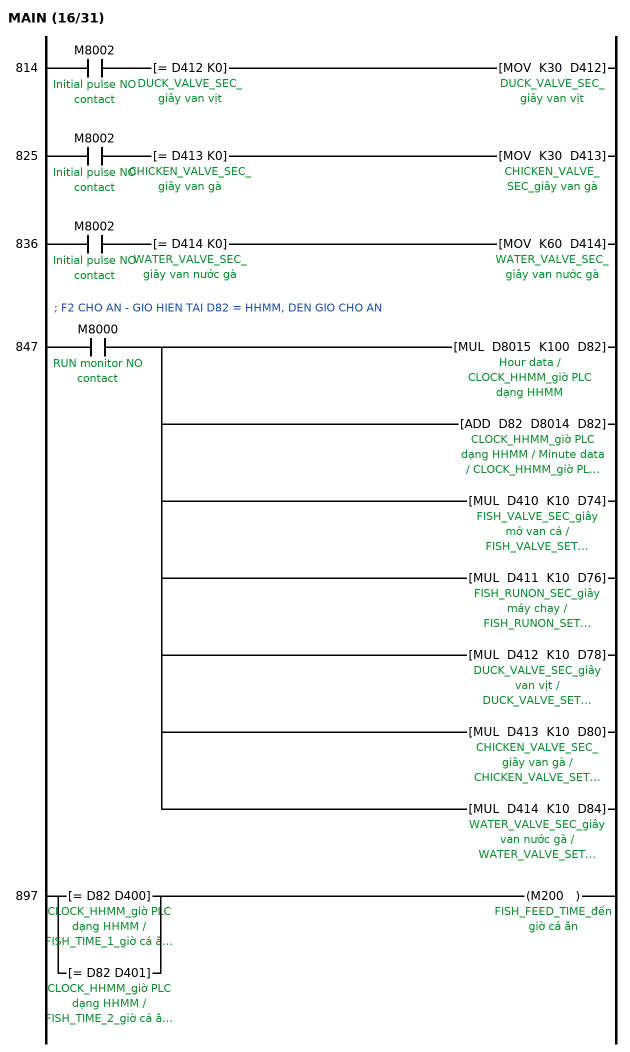
814   LD      M8002  ; Initial pulse NO contact
      AND=    D412 K0  ; DUCK_VALVE_SEC_giây van vịt
      MOV     K30 D412
825   LD      M8002  ; Initial pulse NO contact
      AND=    D413 K0  ; CHICKEN_VALVE_SEC_giây van gà
      MOV     K30 D413
836   LD      M8002  ; Initial pulse NO contact
      AND=    D414 K0  ; WATER_VALVE_SEC_giây van nước gà
      MOV     K60 D414
; F2 CHO AN - GIO HIEN TAI D82 = HHMM, DEN GIO CHO AN
847   LD      M8000  ; RUN monitor NO contact
      MUL     D8015 K100 D82  ; CLOCK_HHMM_giờ PLC dạng HHMM
      ADD     D82 D8014 D82
      MUL     D410 K10 D74  ; FISH_VALVE_SET_D410x10
      MUL     D411 K10 D76  ; FISH_RUNON_SET_D411x10
      MUL     D412 K10 D78  ; DUCK_VALVE_SET_D412x10
      MUL     D413 K10 D80  ; CHICKEN_VALVE_SET_D413x10
      MUL     D414 K10 D84  ; WATER_VALVE_SET_D414x10
897   LD=     D82 D400  ; CLOCK_HHMM_giờ PLC dạng HHMM / FISH_TIME_1_giờ cá ăn 1 HHMM
      OR=     D82 D401  ; CLOCK_HHMM_giờ PLC dạng HHMM / FISH_TIME_2_giờ cá ăn 2 HHMM
      OUT     M200  ; FISH_FEED_TIME_đến giờ cá ăn
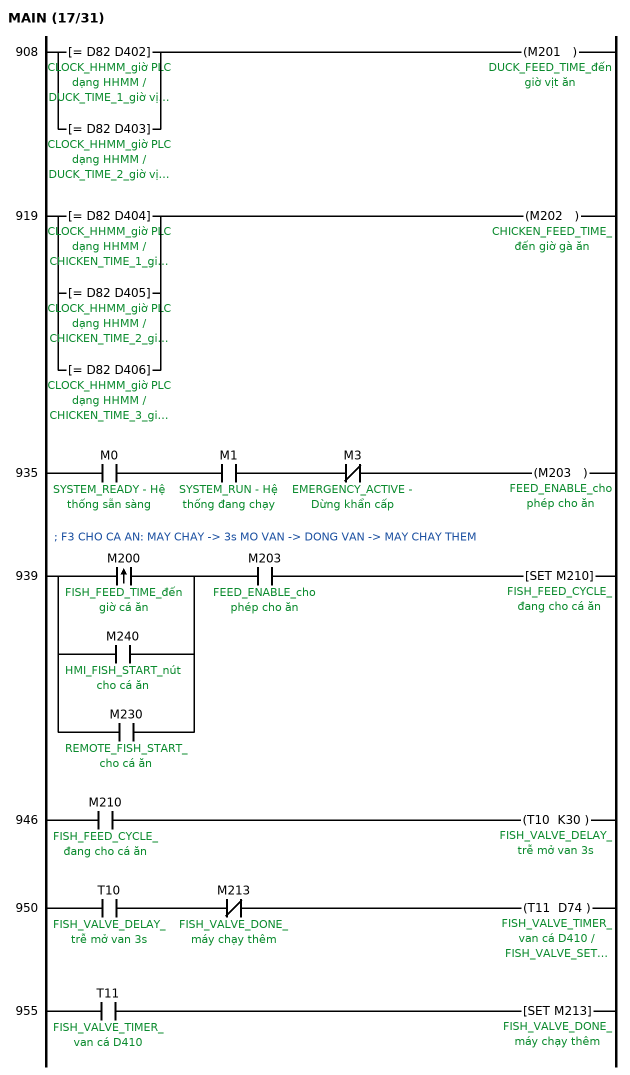
908   LD=     D82 D402  ; CLOCK_HHMM_giờ PLC dạng HHMM / DUCK_TIME_1_giờ vịt ăn 1 HHMM
      OR=     D82 D403  ; CLOCK_HHMM_giờ PLC dạng HHMM / DUCK_TIME_2_giờ vịt ăn 2 HHMM
      OUT     M201  ; DUCK_FEED_TIME_đến giờ vịt ăn
919   LD=     D82 D404  ; CLOCK_HHMM_giờ PLC dạng HHMM / CHICKEN_TIME_1_giờ gà 1 HHMM
      OR=     D82 D405  ; CLOCK_HHMM_giờ PLC dạng HHMM / CHICKEN_TIME_2_giờ gà 2 HHMM
      OR=     D82 D406  ; CLOCK_HHMM_giờ PLC dạng HHMM / CHICKEN_TIME_3_giờ gà 3 HHMM
      OUT     M202  ; CHICKEN_FEED_TIME_đến giờ gà ăn
935   LD      M0  ; SYSTEM_READY - Hệ thống sẵn sàng
      AND     M1  ; SYSTEM_RUN - Hệ thống đang chạy
      ANI     M3  ; EMERGENCY_ACTIVE - Dừng khẩn cấp
      OUT     M203  ; FEED_ENABLE_cho phép cho ăn
; F3 CHO CA AN: MAY CHAY -> 3s MO VAN -> DONG VAN -> MAY CHAY THEM
939   LDP     M200  ; FISH_FEED_TIME_đến giờ cá ăn
      LD      M240  ; HMI_FISH_START_nút cho cá ăn
      OR      M230  ; REMOTE_FISH_START_cho cá ăn
      ORB
      AND     M203  ; FEED_ENABLE_cho phép cho ăn
      SET     M210  ; FISH_FEED_CYCLE_đang cho cá ăn
946   LD      M210  ; FISH_FEED_CYCLE_đang cho cá ăn
      OUT     T10 K30  ; FISH_VALVE_DELAY_trễ mở van 3s
950   LD      T10  ; FISH_VALVE_DELAY_trễ mở van 3s
      ANI     M213  ; FISH_VALVE_DONE_máy chạy thêm
      OUT     T11 D74  ; FISH_VALVE_TIMER_van cá D410 / FISH_VALVE_SET_D410x10
955   LD      T11  ; FISH_VALVE_TIMER_van cá D410
      SET     M213  ; FISH_VALVE_DONE_máy chạy thêm
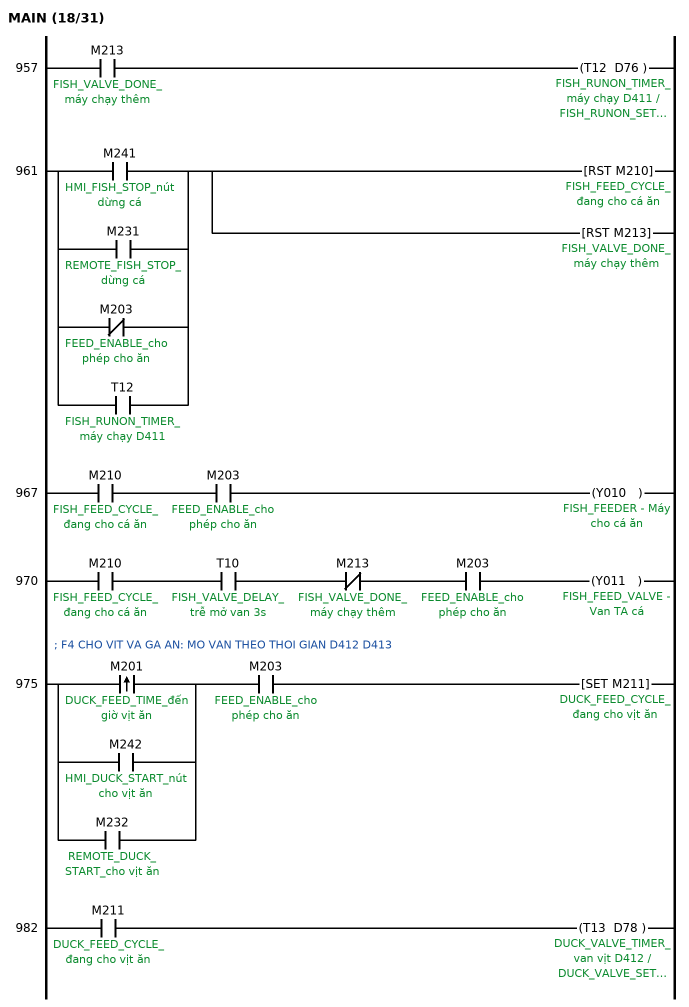
957   LD      M213  ; FISH_VALVE_DONE_máy chạy thêm
      OUT     T12 D76  ; FISH_RUNON_TIMER_máy chạy D411 / FISH_RUNON_SET_D411x10
961   LD      M241  ; HMI_FISH_STOP_nút dừng cá
      OR      M231  ; REMOTE_FISH_STOP_dừng cá
      ORI     M203  ; FEED_ENABLE_cho phép cho ăn
      OR      T12  ; FISH_RUNON_TIMER_máy chạy D411
      RST     M210  ; FISH_FEED_CYCLE_đang cho cá ăn
      RST     M213  ; FISH_VALVE_DONE_máy chạy thêm
967   LD      M210  ; FISH_FEED_CYCLE_đang cho cá ăn
      AND     M203  ; FEED_ENABLE_cho phép cho ăn
      OUT     Y010  ; FISH_FEEDER - Máy cho cá ăn
970   LD      M210  ; FISH_FEED_CYCLE_đang cho cá ăn
      AND     T10  ; FISH_VALVE_DELAY_trễ mở van 3s
      ANI     M213  ; FISH_VALVE_DONE_máy chạy thêm
      AND     M203  ; FEED_ENABLE_cho phép cho ăn
      OUT     Y011  ; FISH_FEED_VALVE - Van TA cá
; F4 CHO VIT VA GA AN: MO VAN THEO THOI GIAN D412 D413
975   LDP     M201  ; DUCK_FEED_TIME_đến giờ vịt ăn
      LD      M242  ; HMI_DUCK_START_nút cho vịt ăn
      OR      M232  ; REMOTE_DUCK_START_cho vịt ăn
      ORB
      AND     M203  ; FEED_ENABLE_cho phép cho ăn
      SET     M211  ; DUCK_FEED_CYCLE_đang cho vịt ăn
982   LD      M211  ; DUCK_FEED_CYCLE_đang cho vịt ăn
      OUT     T13 D78  ; DUCK_VALVE_TIMER_van vịt D412 / DUCK_VALVE_SET_D412x10
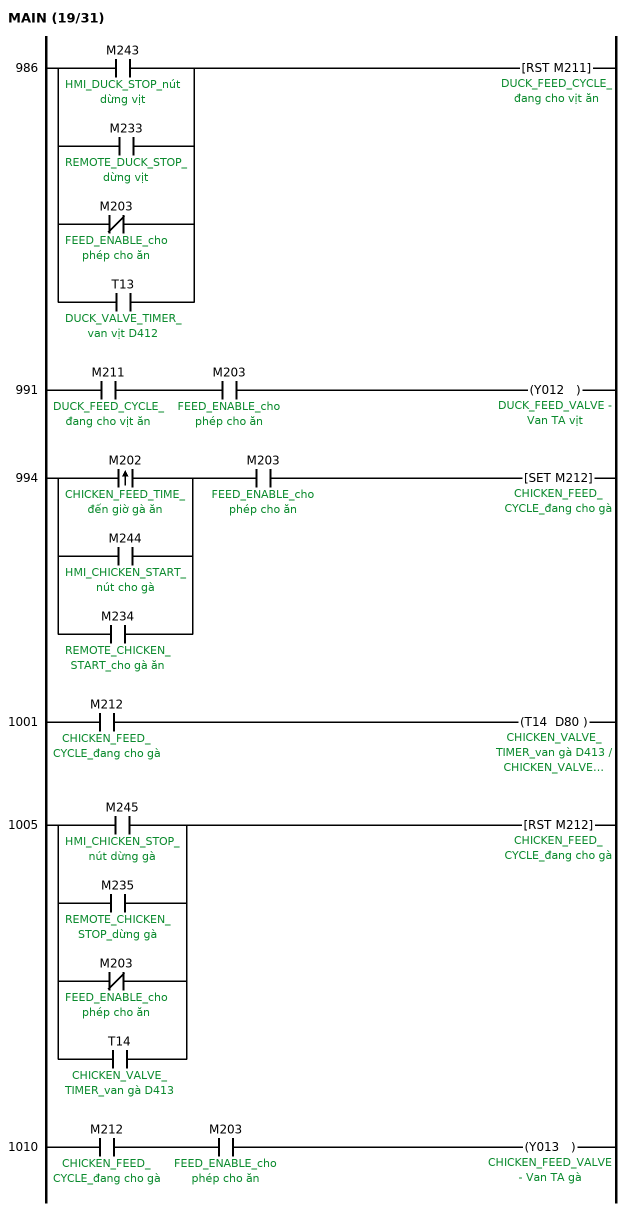
986   LD      M243  ; HMI_DUCK_STOP_nút dừng vịt
      OR      M233  ; REMOTE_DUCK_STOP_dừng vịt
      ORI     M203  ; FEED_ENABLE_cho phép cho ăn
      OR      T13  ; DUCK_VALVE_TIMER_van vịt D412
      RST     M211  ; DUCK_FEED_CYCLE_đang cho vịt ăn
991   LD      M211  ; DUCK_FEED_CYCLE_đang cho vịt ăn
      AND     M203  ; FEED_ENABLE_cho phép cho ăn
      OUT     Y012  ; DUCK_FEED_VALVE - Van TA vịt
994   LDP     M202  ; CHICKEN_FEED_TIME_đến giờ gà ăn
      LD      M244  ; HMI_CHICKEN_START_nút cho gà
      OR      M234  ; REMOTE_CHICKEN_START_cho gà ăn
      ORB
      AND     M203  ; FEED_ENABLE_cho phép cho ăn
      SET     M212  ; CHICKEN_FEED_CYCLE_đang cho gà
1001  LD      M212  ; CHICKEN_FEED_CYCLE_đang cho gà
      OUT     T14 D80  ; CHICKEN_VALVE_TIMER_van gà D413 / CHICKEN_VALVE_SET_D413x10
1005  LD      M245  ; HMI_CHICKEN_STOP_nút dừng gà
      OR      M235  ; REMOTE_CHICKEN_STOP_dừng gà
      ORI     M203  ; FEED_ENABLE_cho phép cho ăn
      OR      T14  ; CHICKEN_VALVE_TIMER_van gà D413
      RST     M212  ; CHICKEN_FEED_CYCLE_đang cho gà
1010  LD      M212  ; CHICKEN_FEED_CYCLE_đang cho gà
      AND     M203  ; FEED_ENABLE_cho phép cho ăn
      OUT     Y013  ; CHICKEN_FEED_VALVE - Van TA gà
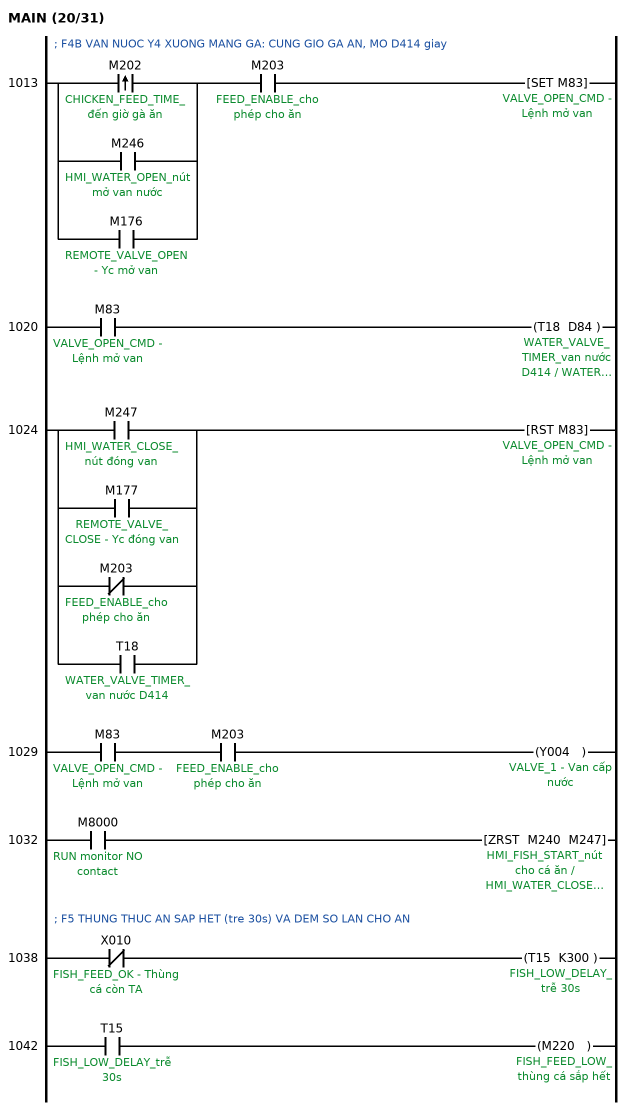
; F4B VAN NUOC Y4 XUONG MANG GA: CUNG GIO GA AN, MO D414 giay
1013  LDP     M202  ; CHICKEN_FEED_TIME_đến giờ gà ăn
      LD      M246  ; HMI_WATER_OPEN_nút mở van nước
      OR      M176  ; REMOTE_VALVE_OPEN - Yc mở van
      ORB
      AND     M203  ; FEED_ENABLE_cho phép cho ăn
      SET     M83  ; VALVE_OPEN_CMD - Lệnh mở van
1020  LD      M83  ; VALVE_OPEN_CMD - Lệnh mở van
      OUT     T18 D84  ; WATER_VALVE_TIMER_van nước D414 / WATER_VALVE_SET_D414x10
1024  LD      M247  ; HMI_WATER_CLOSE_nút đóng van
      OR      M177  ; REMOTE_VALVE_CLOSE - Yc đóng van
      ORI     M203  ; FEED_ENABLE_cho phép cho ăn
      OR      T18  ; WATER_VALVE_TIMER_van nước D414
      RST     M83  ; VALVE_OPEN_CMD - Lệnh mở van
1029  LD      M83  ; VALVE_OPEN_CMD - Lệnh mở van
      AND     M203  ; FEED_ENABLE_cho phép cho ăn
      OUT     Y004  ; VALVE_1 - Van cấp nước
1032  LD      M8000  ; RUN monitor NO contact
      ZRST    M240 M247
; F5 THUNG THUC AN SAP HET (tre 30s) VA DEM SO LAN CHO AN
1038  LDI     X010  ; FISH_FEED_OK - Thùng cá còn TA
      OUT     T15 K300  ; FISH_LOW_DELAY_trễ 30s
1042  LD      T15  ; FISH_LOW_DELAY_trễ 30s
      OUT     M220  ; FISH_FEED_LOW_thùng cá sắp hết
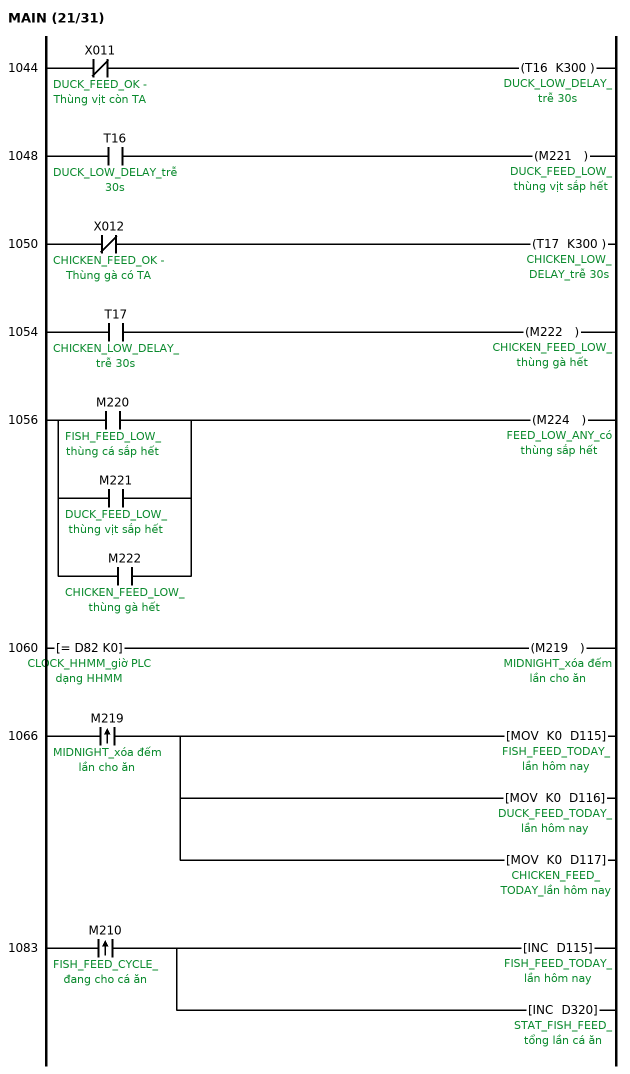
1044  LDI     X011  ; DUCK_FEED_OK - Thùng vịt còn TA
      OUT     T16 K300  ; DUCK_LOW_DELAY_trễ 30s
1048  LD      T16  ; DUCK_LOW_DELAY_trễ 30s
      OUT     M221  ; DUCK_FEED_LOW_thùng vịt sắp hết
1050  LDI     X012  ; CHICKEN_FEED_OK - Thùng gà có TA
      OUT     T17 K300  ; CHICKEN_LOW_DELAY_trễ 30s
1054  LD      T17  ; CHICKEN_LOW_DELAY_trễ 30s
      OUT     M222  ; CHICKEN_FEED_LOW_thùng gà hết
1056  LD      M220  ; FISH_FEED_LOW_thùng cá sắp hết
      OR      M221  ; DUCK_FEED_LOW_thùng vịt sắp hết
      OR      M222  ; CHICKEN_FEED_LOW_thùng gà hết
      OUT     M224  ; FEED_LOW_ANY_có thùng sắp hết
1060  LD=     D82 K0  ; CLOCK_HHMM_giờ PLC dạng HHMM
      OUT     M219  ; MIDNIGHT_xóa đếm lần cho ăn
1066  LDP     M219  ; MIDNIGHT_xóa đếm lần cho ăn
      MOV     K0 D115  ; FISH_FEED_TODAY_lần hôm nay
      MOV     K0 D116  ; DUCK_FEED_TODAY_lần hôm nay
      MOV     K0 D117  ; CHICKEN_FEED_TODAY_lần hôm nay
1083  LDP     M210  ; FISH_FEED_CYCLE_đang cho cá ăn
      INC     D115
      INC     D320  ; STAT_FISH_FEED_tổng lần cá ăn
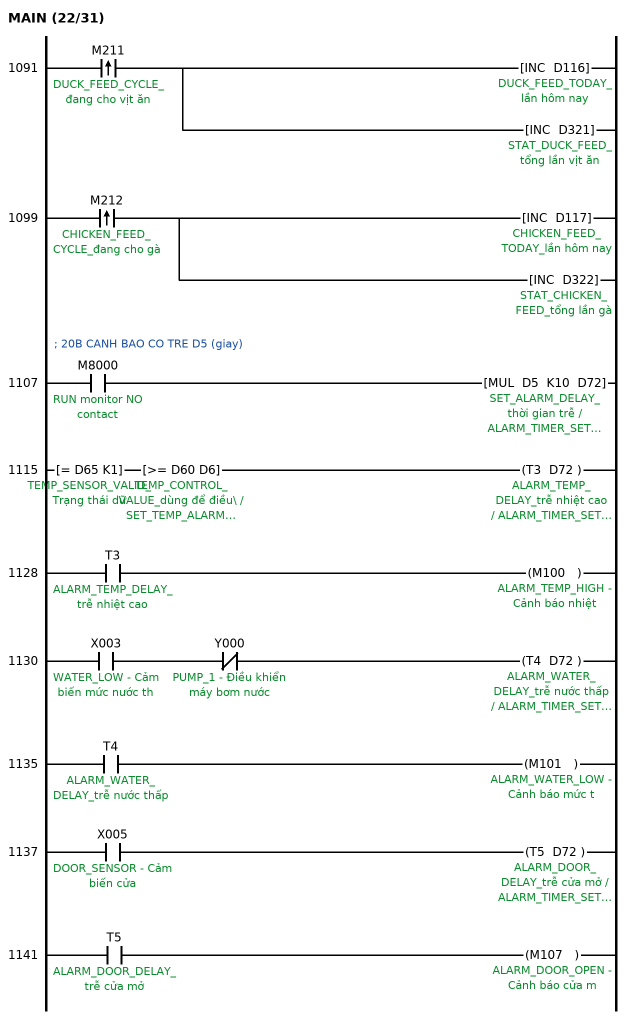
1091  LDP     M211  ; DUCK_FEED_CYCLE_đang cho vịt ăn
      INC     D116
      INC     D321  ; STAT_DUCK_FEED_tổng lần vịt ăn
1099  LDP     M212  ; CHICKEN_FEED_CYCLE_đang cho gà
      INC     D117
      INC     D322  ; STAT_CHICKEN_FEED_tổng lần gà
; 20B CANH BAO CO TRE D5 (giay)
1107  LD      M8000  ; RUN monitor NO contact
      MUL     D5 K10 D72  ; ALARM_TIMER_SET_đặt T3-T5=D5x10
1115  LD=     D65 K1  ; TEMP_SENSOR_VALID_Trạng thái dữ
      AND>=   D60 D6  ; TEMP_CONTROL_VALUE_dùng để điều\ / SET_TEMP_ALARM_HIGH_nhiệt độ cao
      OUT     T3 D72  ; ALARM_TEMP_DELAY_trễ nhiệt cao / ALARM_TIMER_SET_đặt T3-T5=D5x10
1128  LD      T3  ; ALARM_TEMP_DELAY_trễ nhiệt cao
      OUT     M100  ; ALARM_TEMP_HIGH - Cảnh báo nhiệt
1130  LD      X003  ; WATER_LOW - Cảm biến mức nước th
      ANI     Y000  ; PUMP_1 - Điều khiển máy bơm nước
      OUT     T4 D72  ; ALARM_WATER_DELAY_trễ nước thấp / ALARM_TIMER_SET_đặt T3-T5=D5x10
1135  LD      T4  ; ALARM_WATER_DELAY_trễ nước thấp
      OUT     M101  ; ALARM_WATER_LOW - Cảnh báo mức t
1137  LD      X005  ; DOOR_SENSOR - Cảm biến cửa
      OUT     T5 D72  ; ALARM_DOOR_DELAY_trễ cửa mở / ALARM_TIMER_SET_đặt T3-T5=D5x10
1141  LD      T5  ; ALARM_DOOR_DELAY_trễ cửa mở
      OUT     M107  ; ALARM_DOOR_OPEN - Cảnh báo cửa m
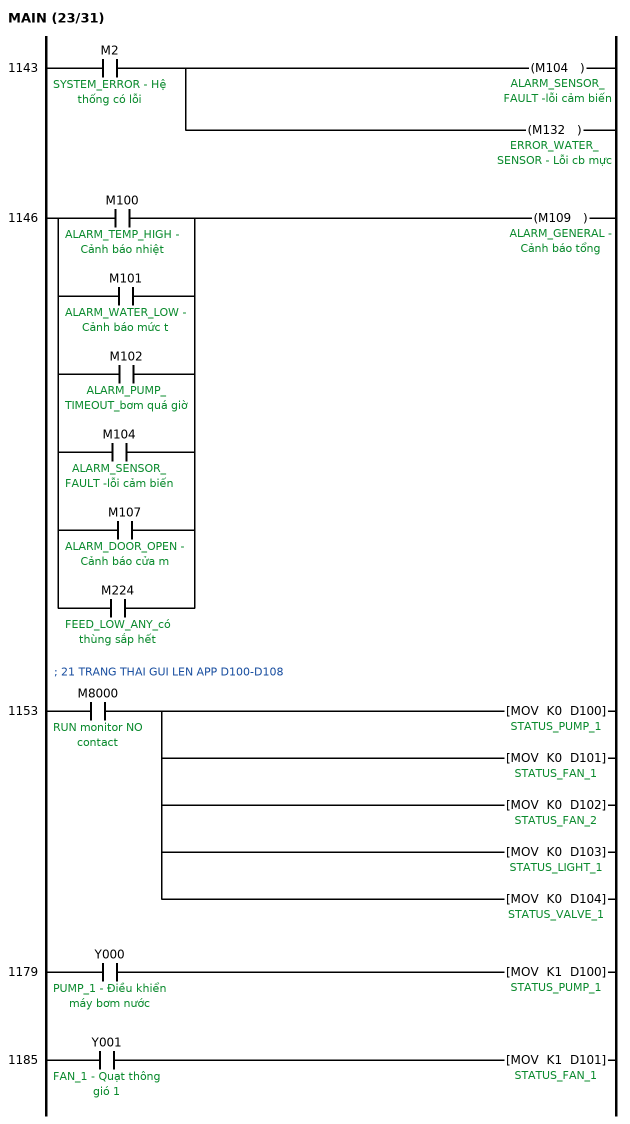
1143  LD      M2  ; SYSTEM_ERROR - Hệ thống có lỗi
      OUT     M104  ; ALARM_SENSOR_FAULT -lỗi cảm biến
      OUT     M132  ; ERROR_WATER_SENSOR - Lỗi cb mực
1146  LD      M100  ; ALARM_TEMP_HIGH - Cảnh báo nhiệt
      OR      M101  ; ALARM_WATER_LOW - Cảnh báo mức t
      OR      M102  ; ALARM_PUMP_TIMEOUT_bơm quá giờ
      OR      M104  ; ALARM_SENSOR_FAULT -lỗi cảm biến
      OR      M107  ; ALARM_DOOR_OPEN - Cảnh báo cửa m
      OR      M224  ; FEED_LOW_ANY_có thùng sắp hết
      OUT     M109  ; ALARM_GENERAL - Cảnh báo tổng
; 21 TRANG THAI GUI LEN APP D100-D108
1153  LD      M8000  ; RUN monitor NO contact
      MOV     K0 D100  ; STATUS_PUMP_1
      MOV     K0 D101  ; STATUS_FAN_1
      MOV     K0 D102  ; STATUS_FAN_2
      MOV     K0 D103  ; STATUS_LIGHT_1
      MOV     K0 D104  ; STATUS_VALVE_1
1179  LD      Y000  ; PUMP_1 - Điều khiển máy bơm nước
      MOV     K1 D100
1185  LD      Y001  ; FAN_1 - Quạt thông gió 1
      MOV     K1 D101
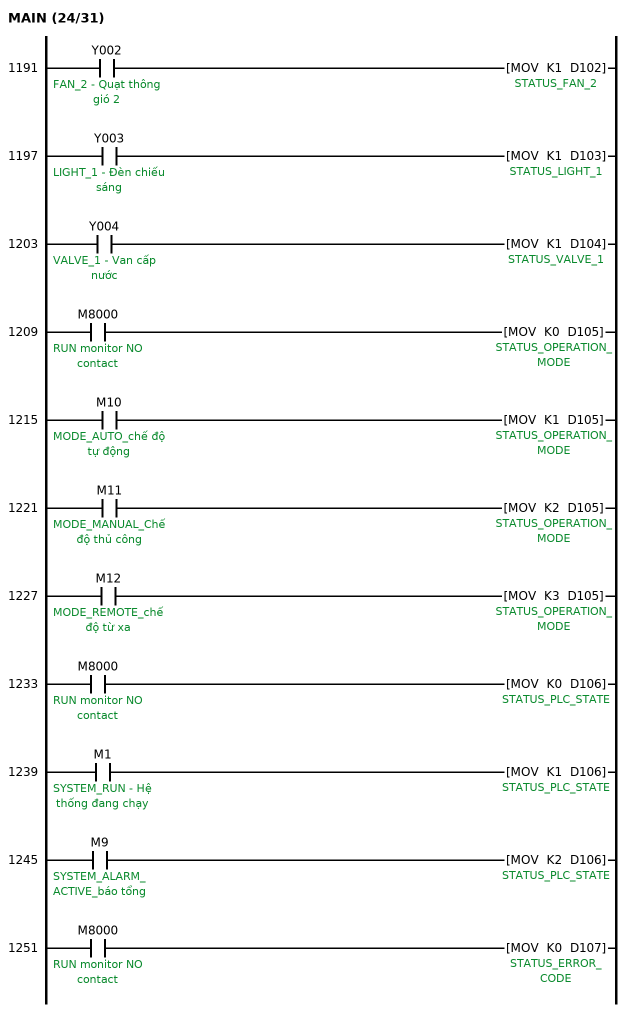
1191  LD      Y002  ; FAN_2 - Quạt thông gió 2
      MOV     K1 D102
1197  LD      Y003  ; LIGHT_1 - Đèn chiếu sáng
      MOV     K1 D103
1203  LD      Y004  ; VALVE_1 - Van cấp nước
      MOV     K1 D104
1209  LD      M8000  ; RUN monitor NO contact
      MOV     K0 D105  ; STATUS_OPERATION_MODE
1215  LD      M10  ; MODE_AUTO_chế độ tự động
      MOV     K1 D105
1221  LD      M11  ; MODE_MANUAL_Chế độ thủ công
      MOV     K2 D105
1227  LD      M12  ; MODE_REMOTE_chế độ từ xa
      MOV     K3 D105
1233  LD      M8000  ; RUN monitor NO contact
      MOV     K0 D106  ; STATUS_PLC_STATE
1239  LD      M1  ; SYSTEM_RUN - Hệ thống đang chạy
      MOV     K1 D106
1245  LD      M9  ; SYSTEM_ALARM_ACTIVE_báo tổng
      MOV     K2 D106
1251  LD      M8000  ; RUN monitor NO contact
      MOV     K0 D107  ; STATUS_ERROR_CODE
